(* IEC 61131-3 sources: avi-aoi-management/scripts/ai-eval/ngau-nhien/kho/st-ud6-nhiet-on-off/khung/src, 2 files *)

(* ---- DieuKhienNhietLo.st ---- *)
FUNCTION_BLOCK DieuKhienNhietLo
VAR_INPUT
    BAT : BOOL;
    NHIET : REAL;
    SP : REAL;
    TRE : REAL;
    NGUONG_CAO : REAL;
    NGUONG_HH : REAL;
    RESET : BOOL;
END_VAR
VAR_OUTPUT
    SUOI : BOOL;
    CANH_BAO_CAO : BOOL;
    NGAT_HH : BOOL;
    LOI_CAM_BIEN : BOOL;
    TRANG_THAI : INT;
END_VAR
    (* TODO: cài đặt theo đề bài *)
    SUOI := FALSE;
END_FUNCTION_BLOCK

(* ---- TreHaiNguong.st ---- *)
FUNCTION_BLOCK TreHaiNguong
VAR_INPUT
    X : REAL;
    SP : REAL;
    TRE : REAL;
END_VAR
VAR_OUTPUT
    Q : BOOL;
END_VAR
    (* TODO: cài đặt theo đề bài *)
    Q := FALSE;
END_FUNCTION_BLOCK
